{region 'Documentation'}
(*!
<summary>Checks calendar-day identity and range bounds despite hidden time-of-day components.</summary>
<description>
Named rows separate independent comparisons by a disabled reset call.
Only explicitly marked escalation rows retain the preceding subject result.
Outer Assertions latch every observation before advancing to the next row.
Intentional findings remain in the local capture; no production algorithm is copied.
</description>
*)
{endregion}
FUNCTION_BLOCK Test_AssertionDateNormalization EXTENDS TestCaseBase
VAR
    FEqualSubject : AssertEqual_Date;
    FInTimespanSubject : AssertInTimespan_Date;
    FNotInTimespanSubject : AssertNotInTimespan_Date;
    FActual : DATE;
    FReference : DATE;
    FStart : DATE;
    FEnd : DATE;
    FExpectedEqualResult : E_Result;
    FExpectedInTimespanResult : E_Result;
    FExpectedNotInTimespanResult : E_Result;
    FExpectedFindings : UDINT;
    FCapture : EventBuffer;
    FEvents : ARRAY[1..CaptureLength] OF ST_Event;
    FCaptureFifo : ST_FifoStatus;
    FCaptureStatus : ST_EventBufferStatus;
    FRow : UINT;
    FRowPrepared : BOOL;
    FPreserveResults : BOOL;
    FObservationReady : BOOL;
    FChecked : BOOL;
    FSetupValid : BOOL;
END_VAR
VAR
    FEqualResult : AssertTrue;
    FEqualResultMatches : BOOL;
    FInTimespanResult : AssertTrue;
    FInTimespanResultMatches : BOOL;
    FNotInTimespanResult : AssertTrue;
    FNotInTimespanResultMatches : BOOL;
    FCaptureIntegrity : AssertTrue;
    FCaptureIntegrityMatches : BOOL;
END_VAR
VAR CONSTANT
    CaptureLength : UINT := 8;
    SameDay : UINT := 1;
    NextDay : UINT := 2;
    NormalizedEqualBounds : UINT := 3;
    ReversedDays : UINT := 4;
    LastRow : UINT := ReversedDays;

END_VAR

SUPER^();

{region 'Documentation'}
(*!
<summary>Collects only outer checking Assertions, never intentional subject findings.</summary>
*)
{endregion}
METHOD PROTECTED AggregateResults
VAR_INPUT
    Aggregator : I_ResultAggregator; //! Borrowed result sink owned by the outer Test Case; add this test's checking Assertions without resetting or retaining the sink.
END_VAR
Aggregator.AddProvider(Provider := FEqualResult);
Aggregator.AddProvider(Provider := FInTimespanResult);
Aggregator.AddProvider(Provider := FNotInTimespanResult);
Aggregator.AddProvider(Provider := FCaptureIntegrity);
END_METHOD

{region 'Documentation'}
(*!
<summary>Calls each inherited production Assertion once using the selected row.</summary>
*)
{endregion}
METHOD PRIVATE CallSubjects
VAR_INPUT
    Enable : BOOL; //! Observation-enable input forwarded to the controlled Assertion subjects for this call.
END_VAR
FEqualSubject(Enable := Enable,
    State := E_State.Running,
    IN := FActual,
    Expected := FReference);
FInTimespanSubject(Enable := Enable,
    State := E_State.Running,
    IN := FActual,
    StartTime := FStart,
    EndTime := FEnd);
FNotInTimespanSubject(Enable := Enable,
    State := E_State.Running,
    IN := FActual,
    StartTime := FStart,
    EndTime := FEnd);
END_METHOD

{region 'Documentation'}
(*!
<summary>Extends base validation with subject and checking-Assertion setup.</summary>
*)
{endregion}
METHOD PROTECTED CheckInitialization : BOOL //! TRUE when the inherited initialization check and this concrete fixture check both accept the setup.
CheckInitialization := SUPER^.CheckInitialization();
IF NOT CheckInitialization THEN
    RETURN;
END_IF;

CheckInitialization := FSetupValid
    AND FEqualResult.IsInitialized
    AND FInTimespanResult.IsInitialized
    AND FNotInTimespanResult.IsInitialized
    AND FCaptureIntegrity.IsInitialized;
IF NOT CheckInitialization THEN
    EventPublisher.PublishEvent(Event := CreateFrameworkEvent(Name := Name,
        ResourceName := '',
        State := State,
        Severity := E_EventSeverity.Error,
        Message := 'Comparison selftest setup failed.'));
END_IF;
END_METHOD

{region 'Documentation'}
(*!
<summary>Checks results and isolated findings against explicit expectations.</summary>
*)
{endregion}
METHOD PRIVATE CheckResults
FEqualResultMatches := FEqualSubject.Result = FExpectedEqualResult;
FInTimespanResultMatches := FInTimespanSubject.Result = FExpectedInTimespanResult;
FNotInTimespanResultMatches := FNotInTimespanSubject.Result = FExpectedNotInTimespanResult;
FCaptureIntegrityMatches := (FCaptureStatus.SequenceId = FExpectedFindings)
    AND (FCaptureStatus.LostEventCount = 0);
END_METHOD

{region 'Documentation'}
(*!
<summary>Configures checking Assertions; subject actions remain in the test script.</summary>
*)
{endregion}
METHOD PROTECTED Configure
VAR
    Initialized : BOOL;
END_VAR
FPreparationStateCount := 0;
FTestStateCount := 1;
FEqualResult.Initialize(Parent := THIS^,
    AssertionName := 'EqualResult');
FInTimespanResult.Initialize(Parent := THIS^,
    AssertionName := 'InTimespanResult');
FNotInTimespanResult.Initialize(Parent := THIS^,
    AssertionName := 'NotInTimespanResult');
FCaptureIntegrity.Initialize(Parent := THIS^,
    AssertionName := 'CaptureIntegrity');
FSetupValid := FCapture.Initialize(Buffer := FEvents,
    FifoControl := FCaptureFifo,
    Status := FCaptureStatus);
FEqualSubject.BindPublisher(Publisher := FCapture);
Initialized := FEqualSubject.Initialize(Parent := THIS^,
    AssertionName := 'EqualSubject');
FSetupValid := FSetupValid AND Initialized;
FInTimespanSubject.BindPublisher(Publisher := FCapture);
Initialized := FInTimespanSubject.Initialize(Parent := THIS^,
    AssertionName := 'InTimespanSubject');
FSetupValid := FSetupValid AND Initialized;
FNotInTimespanSubject.BindPublisher(Publisher := FCapture);
Initialized := FNotInTimespanSubject.Initialize(Parent := THIS^,
    AssertionName := 'NotInTimespanSubject');
FSetupValid := FSetupValid AND Initialized;
END_METHOD

{region 'Documentation'}
(*!
<summary>Completes abort without asynchronous resources.</summary>
*)
{endregion}
METHOD PROTECTED ProcessAbort
VAR_INPUT
    Enable : BOOL; //! Phase permission supplied by the owning Test Case; FALSE does not authorize progression, while observation may continue.
END_VAR
IF Enable THEN
    CompleteAbort();
END_IF;
END_METHOD

{region 'Documentation'}
(*!
<summary>Latches checked observations before the next script step may proceed.</summary>
*)
{endregion}
METHOD PROTECTED ProcessAssertions
VAR_INPUT
    Enable : BOOL; //! Phase permission supplied by the owning Test Case; FALSE does not authorize progression, while observation may continue.
END_VAR
VAR
    Evaluate : BOOL;
END_VAR
Evaluate := Enable AND FObservationReady;
FEqualResult(Enable := Evaluate,
    State := State,
    IN := FEqualResultMatches);
FInTimespanResult(Enable := Evaluate,
    State := State,
    IN := FInTimespanResultMatches);
FNotInTimespanResult(Enable := Evaluate,
    State := State,
    IN := FNotInTimespanResultMatches);
FCaptureIntegrity(Enable := Evaluate,
    State := State,
    IN := FCaptureIntegrityMatches);
IF Evaluate THEN
    FChecked := TRUE;
END_IF;
END_METHOD

{region 'Documentation'}
(*!
<summary>No Preparation phase is required.</summary>
*)
{endregion}
METHOD PROTECTED ProcessPreparations
VAR_INPUT
    // SA0033: Required hook; this test has no Preparation phase.
    {attribute 'analysis' := '-33'}
    Enable : BOOL; //! Phase permission supplied by the owning Test Case; FALSE does not authorize progression, while observation may continue.
END_VAR
END_METHOD

{region 'Documentation'}
(*!
<summary>Restarts the script and resets the checking Assertions.</summary>
*)
{endregion}
METHOD PROTECTED ProcessReset
FRow := SameDay;
FRowPrepared := FALSE;
FChecked := FALSE;
FObservationReady := FALSE;
FEqualResult.Reset();
FEqualResultMatches := TRUE;
FInTimespanResult.Reset();
FInTimespanResultMatches := TRUE;
FNotInTimespanResult.Reset();
FNotInTimespanResultMatches := TRUE;
FCaptureIntegrity.Reset();
FCaptureIntegrityMatches := TRUE;
CompleteReset();
END_METHOD

{region 'Documentation'}
(*!
<summary>Advances one bounded script step per active PLC cycle.</summary>
*)
{endregion}
METHOD PROTECTED ProcessTests
VAR_INPUT
    Enable : BOOL; //! Phase permission supplied by the owning Test Case; FALSE does not authorize progression, while observation may continue.
END_VAR
IF NOT Enable THEN
    RETURN;
END_IF;

IF FChecked THEN
    FChecked := FALSE;
    FObservationReady := FALSE;
    IF FRow = LastRow THEN
        CompleteTests();
        RETURN;
    END_IF;
    FRow := FRow + 1;
    FRowPrepared := FALSE;
END_IF;

IF NOT FRowPrepared THEN
    SelectRow();
    FCapture.Reset();
    IF NOT FPreserveResults THEN
        ResetSubjects();
    END_IF;
    CallSubjects(Enable := FALSE);
    FRowPrepared := TRUE;
ELSE
    CallSubjects(Enable := TRUE);
    CheckResults();
    FObservationReady := TRUE;
END_IF;
END_METHOD

{region 'Documentation'}
(*!
<summary>Requests fresh subject results before the next disabled call.</summary>
*)
{endregion}
METHOD PRIVATE ResetSubjects
FEqualSubject.Reset();
FInTimespanSubject.Reset();
FNotInTimespanSubject.Reset();
END_METHOD

{region 'Documentation'}
(*!
<summary>Selects literal expectations; only named escalation rows retain preceding subject results.</summary>
*)
{endregion}
METHOD PRIVATE SelectRow
FPreserveResults := FALSE;
CASE FRow OF
    SameDay:
        FActual := UDINT_TO_DATE(UDINT#172799);
        FReference := UDINT_TO_DATE(UDINT#86400);
        FStart := UDINT_TO_DATE(UDINT#86400);
        FEnd := UDINT_TO_DATE(UDINT#172799);
        FExpectedEqualResult := E_Result.Passed;
        FExpectedInTimespanResult := E_Result.Passed;
        FExpectedNotInTimespanResult := E_Result.Failed;
        FExpectedFindings := 1;
    NextDay:
        FActual := UDINT_TO_DATE(UDINT#172800);
        FReference := UDINT_TO_DATE(UDINT#86400);
        FStart := UDINT_TO_DATE(UDINT#86400);
        FEnd := UDINT_TO_DATE(UDINT#172799);
        FExpectedEqualResult := E_Result.Failed;
        FExpectedInTimespanResult := E_Result.Failed;
        FExpectedNotInTimespanResult := E_Result.Passed;
        FExpectedFindings := 2;
    NormalizedEqualBounds:
        FActual := UDINT_TO_DATE(UDINT#86400);
        FReference := UDINT_TO_DATE(UDINT#172799);
        FStart := UDINT_TO_DATE(UDINT#172799);
        FEnd := UDINT_TO_DATE(UDINT#86400);
        FExpectedEqualResult := E_Result.Passed;
        FExpectedInTimespanResult := E_Result.Passed;
        FExpectedNotInTimespanResult := E_Result.Failed;
        FExpectedFindings := 1;
    ReversedDays:
        FActual := UDINT_TO_DATE(UDINT#86400);
        FReference := UDINT_TO_DATE(UDINT#86400);
        FStart := UDINT_TO_DATE(UDINT#172800);
        FEnd := UDINT_TO_DATE(UDINT#86400);
        FExpectedEqualResult := E_Result.Passed;
        FExpectedInTimespanResult := E_Result.Error;
        FExpectedNotInTimespanResult := E_Result.Error;
        FExpectedFindings := 2;
ELSE
    Error(Message := 'Unknown comparison test row.');
END_CASE;
END_METHOD

END_FUNCTION_BLOCK

(* stored: Version 1.1.0.1
   POU Test_AssertionDateNormalization: Id {93b72b08-f6af-4389-8064-e242dc499a7f}, SpecialFunc None
   Folder Internal: Id {97856330-a2a9-4970-9a98-d21ee93415d1}
   Method AggregateResults: Id {4188ef35-6f7c-40c6-86e2-37ab86dbff69}
   Method CallSubjects: Id {8842ee33-b4ae-4126-8754-c0cb7c011397}
   Method CheckInitialization: Id {e274c221-7beb-42de-b0c8-d81d87812601}
   Method CheckResults: Id {cdbcb433-1e49-4e93-98e8-741c75ac29d5}
   Method Configure: Id {bcef9f9e-5954-41e3-9f86-3d809427ac40}
   Method ProcessAbort: Id {9a0f4980-d874-4938-86a3-4a32adaf1e10}
   Method ProcessAssertions: Id {46a714a7-21ac-418b-937a-dfbd261990e3}
   Method ProcessPreparations: Id {b9c9fce9-fd2e-436d-9b9b-0c17d5e9431e}
   Method ProcessReset: Id {41eac43a-7284-4bf6-985c-dbbd41e259eb}
   Method ProcessTests: Id {1d6c3e43-3f0f-42d9-9bad-dc6927fc3888}
   Method ResetSubjects: Id {e47e4180-0800-4ac5-a04c-a25f1b7ea55e}
   Method SelectRow: Id {55cefc81-4ee8-4e68-acab-583c10f974ce} *)
